{attribute 'pack_mode' := '1'}
TYPE ST_EssPublishData :
STRUCT
	Header		:	ST_MqttHeader;
	Devices		:	ARRAY[0..GVL_PARAM.ESS_COUNT-1] OF ST_EssPublish_V1;
END_STRUCT
END_TYPE

(* stored: Version 1.1.0.1, ProductVersion 3.1.4024.15
   DUT ST_EssPublishData: Id {9ed7870b-46b2-476a-8226-fbcdc13043c2} *)
